Staubli VAL3: CalToolPos6.pgx

public program CalToolPos6(tool& x_tTool)
  local bool l_bStatus
  local pointRs l_pCenter
  local tool l_t4
  local tool l_t3
  local tool l_t2
  local tool l_t1
  local frame l_fFrame
  local num l_nFrameErr
  local bool l_bBool
  local pointRs l_p5
  local pointRs l_p4
  local pointRs l_p3
  local pointRs l_p2
  local pointRs l_p1
  local pointRs l_p6
begin
  l_bStatus=false
  link(l_pCenter,world)
  //计算中心点坐标
  l_p1=db:pTeach1
  l_p2=db:pTeach2
  l_p3=db:pTeach3
  l_p4=db:pTeach4
  l_p5=db:pTeach5
  l_p6=db:pTeach6
  l_p1.trsf.z=0
  l_p2.trsf.z=0
  l_p3.trsf.z=0
  l_p4.trsf.z=0
  l_p5.trsf.z=0
  l_p6.trsf.z=0
  call _CalpCircle(l_p1,l_p2,l_p3,l_pCenter,l_bStatus)
  //计算工具的xyz
  link(l_p4,world)
  link(l_p5,world)
  link(l_p6,world)
  link(l_fFrame,world)
  l_nFrameErr=setFrame(l_p4,l_p5,l_p6,l_fFrame)
  switch l_nFrameErr
    case 0
      l_pCenter.trsf.rx=l_fFrame.trsf.rx
      l_pCenter.trsf.ry=l_fFrame.trsf.ry
      l_pCenter.trsf.rz=l_fFrame.trsf.rz
      x_tTool.trsf=!l_p4.trsf*l_pCenter.trsf
    break
        case -1,-2
      call db:hmiAlert("DeviationIsTooLarge","info")
    break
  endSwitch
  call db:hmiAlert("SaveInTool1","info")
end
